Fanuc KAREL source: KA00160.KL

PROGRAM KA00160
%NOLOCKGROUP
VAR
  SRC: ARRAY[4] OF REAL
  DST: ARRAY[4] OF VECTOR
BEGIN
  DST = SRC
END KA00160
